TYPE ST_HmiHydraulicsStatus :
STRUCT
	bPresent		: BOOL;
	bEnabled		: BOOL;
	bPumpRunning	: BOOL;
	bSuctionRunning	: BOOL;
	bOilPressureOK	: BOOL;
	bError			: BOOL;
END_STRUCT
END_TYPE

(* stored: Version 1.1.0.1, ProductVersion 3.1.4024.15
   DUT ST_HmiHydraulicsStatus: Id {5a687828-8d91-4d18-9ac6-e3246960874f} *)
